TYPE ST_ExampleStationStatus :
STRUCT
	runStep				: E_ExampleStationRunStep := E_ExampleStationRunStep.Idle; //running sequence step
	allOpen				: BOOL; //both actuators at home (open)
	allClosed			: BOOL; //both actuators at work (closed)
	
	job					: ST_ExampleRequest; //job being worked on
	cycleCount			: UDINT; //completed jobs
	lastCycleTime		: TIME; //duration of the last close/hold/open cycle
	jobsRejected		: UDINT; //requests rejected as invalid
	lastRejectText		: T_MaxString; //reason for the last rejection
	commError			: BOOL; //transaction timed out waiting for the software
END_STRUCT
END_TYPE

(* stored: Version 1.1.0.1, ProductVersion 3.1.4024.12
   DUT ST_ExampleStationStatus: Id {bf60c8ff-6c3e-41e1-8b16-b6c19490999a} *)
